(* IEC 61131-3 sources: codesys-framework/txt/application/WeVe IO (library)/Analog Output/FB_AnalogOutput, 2 files *)

(* ---- Output.prop.st ---- *)
PROPERTY Output : Real

// --- BEGIN IMPLEMENTATION ---

// ----------- SET -----------
VAR
END_VAR

// -- BEGIN IMPLEMENTATION SET --
_rSetPoint := Output;

(* ---- SysPar.prop.st ---- *)
PROPERTY SysPar : SC_SystemParametersAnalogOutput

// --- BEGIN IMPLEMENTATION ---

// ----------- SET -----------
VAR
END_VAR

// -- BEGIN IMPLEMENTATION SET --
_scSysPar := SysPar;
